Universal Robots PolyScope program: ManyMoves.urp

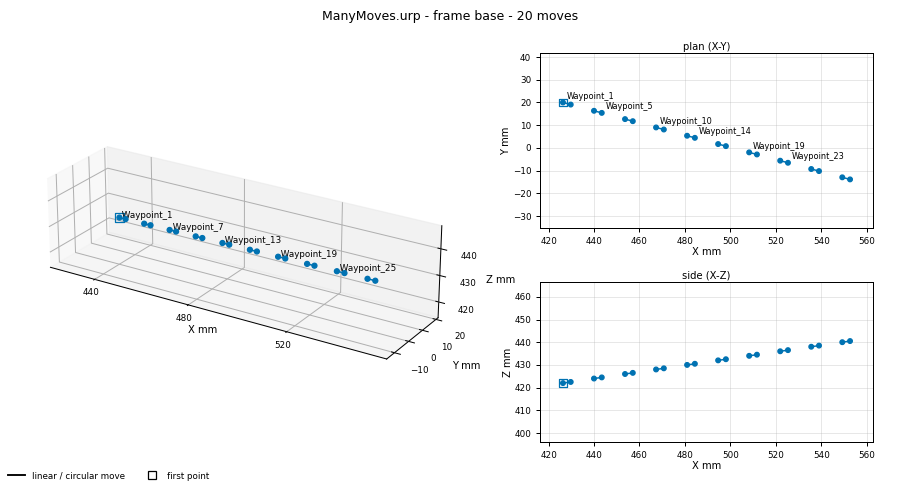
[picture p0: tool path of ManyMoves.urp in frame base, 20 of 30 moves have a stored position in this frame; points joined in program order, loops and branches not executed]
Program ManyMoves (createdIn=3.0.0 lastSavedIn=3.0.0 directory=/programs installation=default)
Robot Program (runOnlyOnce=true motionType=MoveJ speed=1.047198 acceleration=1.396263 useActiveTCP=false)
  'Program generated by RoboDK v6.0.7 for ABB IRB 120-3/0.6 on XX/XX/XXXX 18:00:00'
  'Using nominal kinematics.'
  'Using Ref. Frame S: p[1.234570, -0.098765, 0.050500, 0.000000, 0.000000, 0.523599]'
  'Using TCP Tool S: p[0.010000, 0.020000, 0.150000, 0.000000, 0.000000, 0.000000]'
  Script: set_tcp(p[0.010000, 0.020000, 0.150000, 0.000000, 0.000000, 0.000000])
  Script: movej([0.000000, -0.174533, 0.349066, 0.000000, 0.523599, 0.000000],1.20000,0.75000,0,0.0000)
  MoveJ speed 42.97 deg/s, acceleration 68.75 deg/s^2 (useActiveTCP=true)
    Waypoint Waypoint_1: TCP in base x=426.318 y=20 z=422.034 mm, rx=0.1383 ry=2.2532 rz=-0.2966 rad; joints [0, -10, 20, 0, 30, 0] deg; flange x=317.789 y=39.504 z=526.155 mm, rx=0.1383 ry=2.2532 rz=-0.2966 rad
  MoveL speed 500 mm/s, acceleration 1200 mm/s^2 (useActiveTCP=true)
    Waypoint Waypoint_2: TCP in base x=429.733 y=19.085 z=422.534 mm, rx=0.1383 ry=2.2532 rz=-0.2966 rad; joints [0, -10, 20, 0, 30, 0] deg; flange x=321.204 y=38.589 z=526.655 mm, rx=0.1383 ry=2.2532 rz=-0.2966 rad
  Script: movej([0.349066, -0.174533, 0.349066, 0.000000, 0.523599, 0.000000],1.20000,0.75000,0,0.0000)
  MoveL speed 500 mm/s, acceleration 1200 mm/s^2 (useActiveTCP=true)
    Waypoint Waypoint_3: position(joints=0.000000, -0.174533, 0.349066, 0.000000, 0.523599, 0.000000)
  Script: movej([0.000000, -0.174533, 0.349066, 0.000000, 0.523599, 0.000000],1.20000,0.75000,0,0.0000)
  MoveJ speed 42.97 deg/s, acceleration 68.75 deg/s^2 (useActiveTCP=true)
    Waypoint Waypoint_4: TCP in base x=439.978 y=16.34 z=424.034 mm, rx=0.1383 ry=2.2532 rz=-0.2966 rad; joints [0, -10, 20, 0, 30, 0] deg; flange x=331.449 y=35.844 z=528.155 mm, rx=0.1383 ry=2.2532 rz=-0.2966 rad
  MoveL speed 500 mm/s, acceleration 1200 mm/s^2 (useActiveTCP=true)
    Waypoint Waypoint_5: TCP in base x=443.393 y=15.425 z=424.534 mm, rx=0.1383 ry=2.2532 rz=-0.2966 rad; joints [0, -10, 20, 0, 30, 0] deg; flange x=334.865 y=34.929 z=528.655 mm, rx=0.1383 ry=2.2532 rz=-0.2966 rad
  Script: movej([0.349066, -0.174533, 0.349066, 0.000000, 0.523599, 0.000000],1.20000,0.75000,0,0.0000)
  MoveL speed 500 mm/s, acceleration 1200 mm/s^2 (useActiveTCP=true)
    Waypoint Waypoint_6: position(joints=0.000000, -0.174533, 0.349066, 0.000000, 0.523599, 0.000000)
  Script: movej([0.000000, -0.174533, 0.349066, 0.000000, 0.523599, 0.000000],1.20000,0.75000,0,0.0000)
  MoveJ speed 42.97 deg/s, acceleration 68.75 deg/s^2 (useActiveTCP=true)
    Waypoint Waypoint_7: TCP in base x=453.638 y=12.68 z=426.034 mm, rx=0.1383 ry=2.2532 rz=-0.2966 rad; joints [0, -10, 20, 0, 30, 0] deg; flange x=345.11 y=32.184 z=530.155 mm, rx=0.1383 ry=2.2532 rz=-0.2966 rad
  MoveL speed 500 mm/s, acceleration 1200 mm/s^2 (useActiveTCP=true)
    Waypoint Waypoint_8: TCP in base x=457.054 y=11.765 z=426.534 mm, rx=0.1383 ry=2.2532 rz=-0.2966 rad; joints [0, -10, 20, 0, 30, 0] deg; flange x=348.525 y=31.269 z=530.655 mm, rx=0.1383 ry=2.2532 rz=-0.2966 rad
  Script: movej([0.349066, -0.174533, 0.349066, 0.000000, 0.523599, 0.000000],1.20000,0.75000,0,0.0000)
  MoveL speed 500 mm/s, acceleration 1200 mm/s^2 (useActiveTCP=true)
    Waypoint Waypoint_9: position(joints=0.000000, -0.174533, 0.349066, 0.000000, 0.523599, 0.000000)
  Script: movej([0.000000, -0.174533, 0.349066, 0.000000, 0.523599, 0.000000],1.20000,0.75000,0,0.0000)
  MoveJ speed 42.97 deg/s, acceleration 68.75 deg/s^2 (useActiveTCP=true)
    Waypoint Waypoint_10: TCP in base x=467.299 y=9.019 z=428.034 mm, rx=0.1383 ry=2.2532 rz=-0.2966 rad; joints [0, -10, 20, 0, 30, 0] deg; flange x=358.77 y=28.524 z=532.155 mm, rx=0.1383 ry=2.2532 rz=-0.2966 rad
  MoveL speed 500 mm/s, acceleration 1200 mm/s^2 (useActiveTCP=true)
    Waypoint Waypoint_11: TCP in base x=470.714 y=8.104 z=428.534 mm, rx=0.1383 ry=2.2532 rz=-0.2966 rad; joints [0, -10, 20, 0, 30, 0] deg; flange x=362.185 y=27.609 z=532.655 mm, rx=0.1383 ry=2.2532 rz=-0.2966 rad
  Script: movej([0.349066, -0.174533, 0.349066, 0.000000, 0.523599, 0.000000],1.20000,0.75000,0,0.0000)
  MoveL speed 500 mm/s, acceleration 1200 mm/s^2 (useActiveTCP=true)
    Waypoint Waypoint_12: position(joints=0.000000, -0.174533, 0.349066, 0.000000, 0.523599, 0.000000)
  Script: movej([0.000000, -0.174533, 0.349066, 0.000000, 0.523599, 0.000000],1.20000,0.75000,0,0.0000)
  MoveJ speed 42.97 deg/s, acceleration 68.75 deg/s^2 (useActiveTCP=true)
    Waypoint Waypoint_13: TCP in base x=480.959 y=5.359 z=430.034 mm, rx=0.1383 ry=2.2532 rz=-0.2966 rad; joints [0, -10, 20, 0, 30, 0] deg; flange x=372.43 y=24.863 z=534.155 mm, rx=0.1383 ry=2.2532 rz=-0.2966 rad
  MoveL speed 500 mm/s, acceleration 1200 mm/s^2 (useActiveTCP=true)
    Waypoint Waypoint_14: TCP in base x=484.374 y=4.444 z=430.534 mm, rx=0.1383 ry=2.2532 rz=-0.2966 rad; joints [0, -10, 20, 0, 30, 0] deg; flange x=375.845 y=23.948 z=534.655 mm, rx=0.1383 ry=2.2532 rz=-0.2966 rad
  Script: movej([0.349066, -0.174533, 0.349066, 0.000000, 0.523599, 0.000000],1.20000,0.75000,0,0.0000)
  MoveL speed 500 mm/s, acceleration 1200 mm/s^2 (useActiveTCP=true)
    Waypoint Waypoint_15: position(joints=0.000000, -0.174533, 0.349066, 0.000000, 0.523599, 0.000000)
  Script: movej([0.000000, -0.174533, 0.349066, 0.000000, 0.523599, 0.000000],1.20000,0.75000,0,0.0000)
  MoveJ speed 42.97 deg/s, acceleration 68.75 deg/s^2 (useActiveTCP=true)
    Waypoint Waypoint_16: TCP in base x=494.619 y=1.699 z=432.034 mm, rx=0.1383 ry=2.2532 rz=-0.2966 rad; joints [0, -10, 20, 0, 30, 0] deg; flange x=386.09 y=21.203 z=536.155 mm, rx=0.1383 ry=2.2532 rz=-0.2966 rad
  MoveL speed 500 mm/s, acceleration 1200 mm/s^2 (useActiveTCP=true)
    Waypoint Waypoint_17: TCP in base x=498.034 y=0.784 z=432.534 mm, rx=0.1383 ry=2.2532 rz=-0.2966 rad; joints [0, -10, 20, 0, 30, 0] deg; flange x=389.506 y=20.288 z=536.655 mm, rx=0.1383 ry=2.2532 rz=-0.2966 rad
  Script: movej([0.349066, -0.174533, 0.349066, 0.000000, 0.523599, 0.000000],1.20000,0.75000,0,0.0000)
  MoveL speed 500 mm/s, acceleration 1200 mm/s^2 (useActiveTCP=true)
    Waypoint Waypoint_18: position(joints=0.000000, -0.174533, 0.349066, 0.000000, 0.523599, 0.000000)
  Script: movej([0.000000, -0.174533, 0.349066, 0.000000, 0.523599, 0.000000],1.20000,0.75000,0,0.0000)
  MoveJ speed 42.97 deg/s, acceleration 68.75 deg/s^2 (useActiveTCP=true)
    Waypoint Waypoint_19: TCP in base x=508.28 y=-1.961 z=434.034 mm, rx=0.1383 ry=2.2532 rz=-0.2966 rad; joints [0, -10, 20, 0, 30, 0] deg; flange x=399.751 y=17.543 z=538.155 mm, rx=0.1383 ry=2.2532 rz=-0.2966 rad
  MoveL speed 500 mm/s, acceleration 1200 mm/s^2 (useActiveTCP=true)
    Waypoint Waypoint_20: TCP in base x=511.695 y=-2.876 z=434.534 mm, rx=0.1383 ry=2.2532 rz=-0.2966 rad; joints [0, -10, 20, 0, 30, 0] deg; flange x=403.166 y=16.628 z=538.655 mm, rx=0.1383 ry=2.2532 rz=-0.2966 rad
  Script: movej([0.349066, -0.174533, 0.349066, 0.000000, 0.523599, 0.000000],1.20000,0.75000,0,0.0000)
  MoveL speed 500 mm/s, acceleration 1200 mm/s^2 (useActiveTCP=true)
    Waypoint Waypoint_21: position(joints=0.000000, -0.174533, 0.349066, 0.000000, 0.523599, 0.000000)
  Script: movej([0.000000, -0.174533, 0.349066, 0.000000, 0.523599, 0.000000],1.20000,0.75000,0,0.0000)
  MoveJ speed 42.97 deg/s, acceleration 68.75 deg/s^2 (useActiveTCP=true)
    Waypoint Waypoint_22: TCP in base x=521.94 y=-5.622 z=436.034 mm, rx=0.1383 ry=2.2532 rz=-0.2966 rad; joints [0, -10, 20, 0, 30, 0] deg; flange x=413.411 y=13.883 z=540.155 mm, rx=0.1383 ry=2.2532 rz=-0.2966 rad
  MoveL speed 500 mm/s, acceleration 1200 mm/s^2 (useActiveTCP=true)
    Waypoint Waypoint_23: TCP in base x=525.355 y=-6.537 z=436.534 mm, rx=0.1383 ry=2.2532 rz=-0.2966 rad; joints [0, -10, 20, 0, 30, 0] deg; flange x=416.826 y=12.968 z=540.655 mm, rx=0.1383 ry=2.2532 rz=-0.2966 rad
  Script: movej([0.349066, -0.174533, 0.349066, 0.000000, 0.523599, 0.000000],1.20000,0.75000,0,0.0000)
  MoveL speed 500 mm/s, acceleration 1200 mm/s^2 (useActiveTCP=true)
    Waypoint Waypoint_24: position(joints=0.000000, -0.174533, 0.349066, 0.000000, 0.523599, 0.000000)
  Script: movej([0.000000, -0.174533, 0.349066, 0.000000, 0.523599, 0.000000],1.20000,0.75000,0,0.0000)
  MoveJ speed 42.97 deg/s, acceleration 68.75 deg/s^2 (useActiveTCP=true)
    Waypoint Waypoint_25: TCP in base x=535.6 y=-9.282 z=438.034 mm, rx=0.1383 ry=2.2532 rz=-0.2966 rad; joints [0, -10, 20, 0, 30, 0] deg; flange x=427.071 y=10.222 z=542.155 mm, rx=0.1383 ry=2.2532 rz=-0.2966 rad
  MoveL speed 500 mm/s, acceleration 1200 mm/s^2 (useActiveTCP=true)
    Waypoint Waypoint_26: TCP in base x=539.015 y=-10.197 z=438.534 mm, rx=0.1383 ry=2.2532 rz=-0.2966 rad; joints [0, -10, 20, 0, 30, 0] deg; flange x=430.486 y=9.307 z=542.655 mm, rx=0.1383 ry=2.2532 rz=-0.2966 rad
  Script: movej([0.349066, -0.174533, 0.349066, 0.000000, 0.523599, 0.000000],1.20000,0.75000,0,0.0000)
  MoveL speed 500 mm/s, acceleration 1200 mm/s^2 (useActiveTCP=true)
    Waypoint Waypoint_27: position(joints=0.000000, -0.174533, 0.349066, 0.000000, 0.523599, 0.000000)
  Script: movej([0.000000, -0.174533, 0.349066, 0.000000, 0.523599, 0.000000],1.20000,0.75000,0,0.0000)
  MoveJ speed 42.97 deg/s, acceleration 68.75 deg/s^2 (useActiveTCP=true)
    Waypoint Waypoint_28: TCP in base x=549.26 y=-12.942 z=440.034 mm, rx=0.1383 ry=2.2532 rz=-0.2966 rad; joints [0, -10, 20, 0, 30, 0] deg; flange x=440.731 y=6.562 z=544.155 mm, rx=0.1383 ry=2.2532 rz=-0.2966 rad
  MoveL speed 500 mm/s, acceleration 1200 mm/s^2 (useActiveTCP=true)
    Waypoint Waypoint_29: TCP in base x=552.675 y=-13.857 z=440.534 mm, rx=0.1383 ry=2.2532 rz=-0.2966 rad; joints [0, -10, 20, 0, 30, 0] deg; flange x=444.147 y=5.647 z=544.655 mm, rx=0.1383 ry=2.2532 rz=-0.2966 rad
  Script: movej([0.349066, -0.174533, 0.349066, 0.000000, 0.523599, 0.000000],1.20000,0.75000,0,0.0000)
  MoveL speed 500 mm/s, acceleration 1200 mm/s^2 (useActiveTCP=true)
    Waypoint Waypoint_30: position(joints=0.000000, -0.174533, 0.349066, 0.000000, 0.523599, 0.000000)
